FUNCTION_BLOCK basicValvulaSolenoide (* Valvula solenoide on/off: aberta/fechada pelo fim de curso (se houver) ou pelo comando, e alarme de discrepancia *)
  (* Standard: 61499-2 *)
  (* Version 1.0, 04/11/2026, Hidryco, Hidryco, 1.0: criado para as SV-900 (agua de servico do lodo) *)
  PACKAGE Hidryco.HidrycoLib;
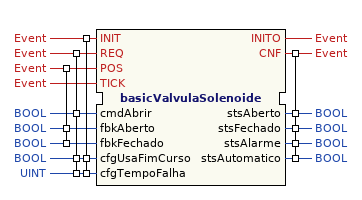
  EVENT_INPUT
    INIT WITH cfgUsaFimCurso, cfgTempoFalha; (* Inicializacao *)
    REQ WITH cmdAbrir, cfgUsaFimCurso, cfgTempoFalha; (* Novo comando da logica *)
    POS WITH fbkAberto, fbkFechado; (* Novo estado dos fins de curso *)
    TICK; (* Base de tempo de 1 s *)
  END_EVENT
  EVENT_OUTPUT
    INITO; (* Inicializacao concluida *)
    CNF WITH stsAberto, stsFechado, stsAlarme, stsAutomatico; (* Estado atualizado *)
  END_EVENT
  VAR_INPUT
    cmdAbrir : BOOL; (* Comando abrir (saida digital da solenoide) *)
    fbkAberto : BOOL; (* Fim de curso aberta (campo) *)
    fbkFechado : BOOL; (* Fim de curso fechada (campo) *)
    cfgUsaFimCurso : BOOL := FALSE; (* TRUE = aberta/fechada pelos fins de curso e alarme de discrepancia; FALSE = pelo comando, sem alarme *)
    cfgTempoFalha : UINT := 10; (* Tempo de discrepancia entre comando e fim de curso para o alarme (s) *)
  END_VAR
  VAR_OUTPUT
    stsAberto : BOOL; (* Valvula aberta *)
    stsFechado : BOOL; (* Valvula fechada *)
    stsAlarme : BOOL; (* Discrepancia entre comando e fim de curso (so com cfgUsaFimCurso) *)
    stsAutomatico : BOOL; (* Sempre FALSE: as SV sao so manuais *)
  END_VAR
  VAR
    discrepancia : BOOL; (* Comando e fim de curso diferentes agora *)
    contagem : UINT; (* Segundos em discrepancia *)
  END_VAR
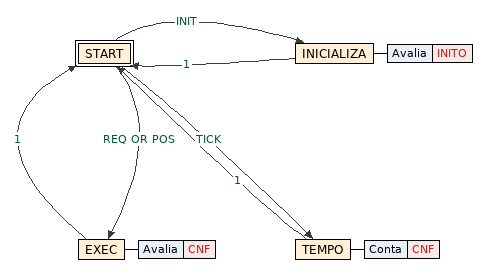
  EC_STATES
    START; (* Initial State *)
    INICIALIZA : Avalia -> INITO;
    EXEC : Avalia -> CNF;
    TEMPO : Conta -> CNF;
  END_STATES
  EC_TRANSITIONS
    START TO INICIALIZA := INIT;
    INICIALIZA TO START := 1;
    START TO EXEC := REQ OR POS;
    EXEC TO START := 1;
    START TO TEMPO := TICK;
    TEMPO TO START := 1;
  END_TRANSITIONS
  ALGORITHM Avalia IN ST: (* Estado pela posicao ou pelo comando *)
IF cfgUsaFimCurso THEN
  stsAberto := fbkAberto;
  stsFechado := fbkFechado;
  discrepancia := (cmdAbrir AND NOT fbkAberto) OR (NOT cmdAbrir AND NOT fbkFechado) OR (fbkAberto AND fbkFechado);
ELSE
  stsAberto := cmdAbrir;
  stsFechado := NOT cmdAbrir;
  discrepancia := FALSE;
END_IF;
IF NOT discrepancia THEN
  contagem := 0;
  stsAlarme := FALSE;
END_IF;
stsAutomatico := FALSE;
  END_ALGORITHM
  ALGORITHM Conta IN ST: (* Conta o tempo de discrepancia (1 s por TICK) *)
IF discrepancia THEN
  IF contagem < 65535 THEN
    contagem := contagem + 1;
  END_IF;
  stsAlarme := contagem >= cfgTempoFalha;
END_IF;
  END_ALGORITHM
END_FUNCTION_BLOCK
